RoboDK station: PickAndPlace(Sriman).rdk

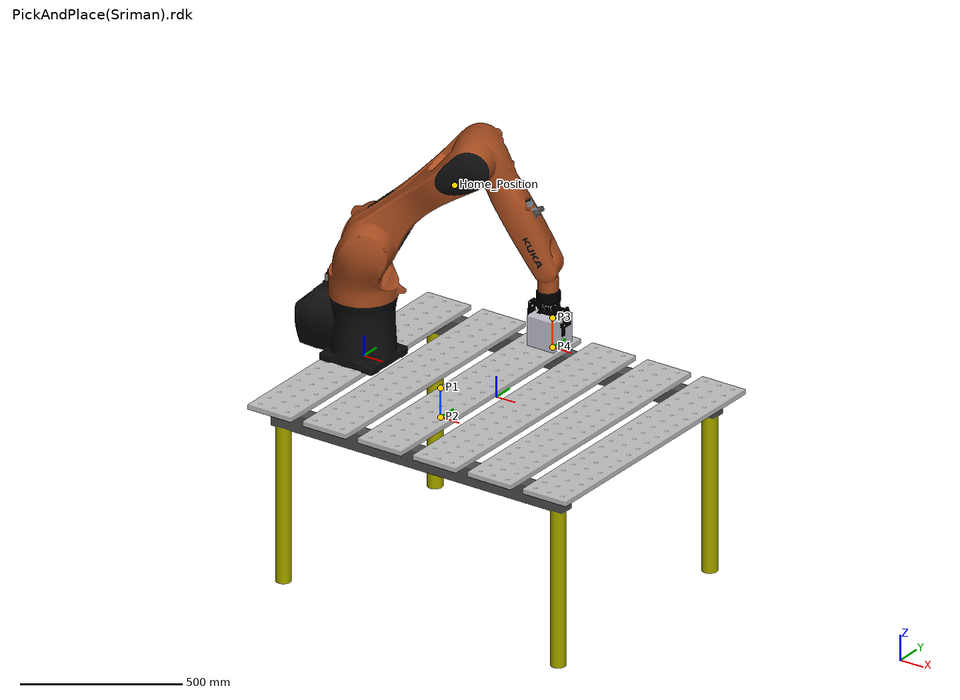
[picture v0: the station drawn from its stored meshes, robots at their saved joint values, targets as dots, program paths as lines]
Station PickAndPlace(Sriman) (saved by RoboDK 6.1.1). Poses are relative to the parent item; angles as X-Y-Z fixed-axis rotations.
  - frame KUKA KR 10 R900 sixx Base at (-500, 0, 0) mm
    - robot KUKA KR 10 R900 sixx: 6 axes, payload 10 kg, reach 901 mm, repeatability 0.03 mm, weight 52 kg
        modified DH rows (alpha deg, a mm, theta deg, d mm): 0, 0, 0, 400; -90, 25, 0, 0; 0, 455, -90, 0; -90, 35, 0, 420; 90, 0, 0, 0; -90, 0, 180, 80
        joint limits [-170, -190, -120, -185, -120, -350] to [170, 45, 156, 185, 120, 350]; home [0, -90, 90, 0, 0, 0]; saved at [-23.826, -44.011, 106.474, 1.623, 26.015, -25.275]
      - tool RobotiQ 2F-85 Gripper (Open), TCP at (0, 0, 130) mm, size 147.4 x 75 x 146.8 mm
        - object box at (0, 0, 0) mm, rotated rx 180 ry -1.8 rz -180 deg, size 100 x 100 x 100 mm, geometry from box.sld
  - frame Base at (0, 0, 0) mm
    - object Table 1200x1000mm (Welding) at (0, 0, 0) mm, size 1193.8 x 965.2 x 609.6 mm, geometry from Table-1200x1000mm-Welding.sld
    - target Home_Position (Cartesian target) at (-158.4, 0, 680.11) mm, rotated rx 180 ry 1.8 rz -180 deg; joints [0, -103.82, 102.02, 0, 90, 0] of KUKA KR 10 R900 sixx
  - frame Pick_Position at (0, -300, 50) mm
    - target P2 (Cartesian target) at (0, 0, 0) mm, rotated rx 180 ry 1.8 rz -180 deg; joints [31.3, -32.692, 103.737, -3.121, 17.441, 34.266] of KUKA KR 10 R900 sixx
    - target P1 (Cartesian target) at (0, 0, 100) mm, rotated rx 180 ry 1.8 rz -180 deg; joints [31.3, -44.011, 106.474, -2.132, 26.015, 33.204] of KUKA KR 10 R900 sixx
  - frame Place_Position at (0, 300, 50) mm
    - target P3 (Cartesian target) at (0, 0, 100) mm, rotated rx 180 ry 1.8 rz -180 deg; joints [-31.3, -44.011, 106.474, 2.132, 26.015, -33.204] of KUKA KR 10 R900 sixx
    - target P4 (Cartesian target) at (0, 0, 0) mm, rotated rx 180 ry 1.8 rz -180 deg; joints [-31.3, -32.692, 103.737, 3.121, 17.441, -34.266] of KUKA KR 10 R900 sixx
  - program Restore (1 instructions, listed below)
  - program Pick (6 instructions, listed below)
  - program Main Program (3 instructions, listed below)
  - program Place (6 instructions, listed below)
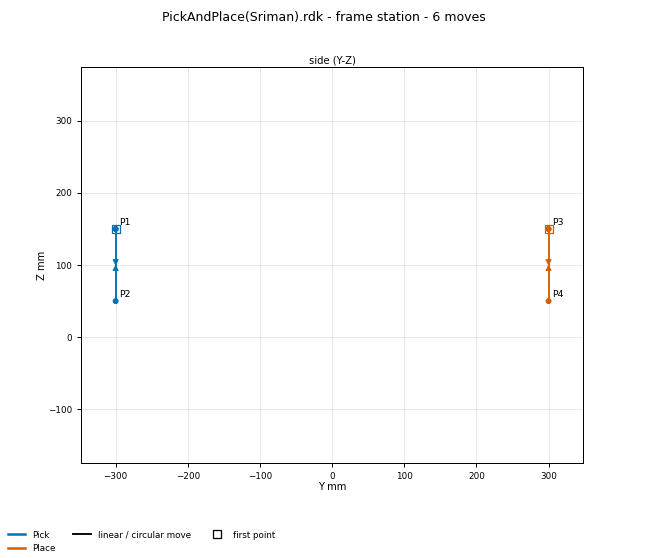
[picture p0: tool path of PickAndPlace(Sriman).rdk in frame station, 6 of 6 moves have a stored position in this frame; points joined in program order, loops and branches not executed]

--- program Restore (robot KUKA KR 10 R900 sixx) ---
  Move objects

--- program Pick (robot KUKA KR 10 R900 sixx) ---
  Set Ref.: Pick_Position
  Set Tool: RobotiQ 2F-85 Gripper (Open)
  MoveJ (P1)
  MoveL (P2)
  Attach to RobotiQ 2F-85 Gripper (Open)
  MoveL (P1)

--- program Main Program (robot KUKA KR 10 R900 sixx) ---
  Call Pick
  Call Place
  Call Restore

--- program Place (robot KUKA KR 10 R900 sixx) ---
  Set Ref.: Place_Position
  Set Tool: RobotiQ 2F-85 Gripper (Open)
  MoveJ (P3)
  MoveL (P4)
  Detach from RobotiQ 2F-85 Gripper (Open)
  MoveL (P3)
